TYPE "ST_CylinderHal"
VERSION : 0.1
   STRUCT
      FeedbackExtended : Bool;
      FeedbackRetracted : Bool;
      ExtendPermit : Bool;
      RetractPermit : Bool;
      PermitDiagnostic : "ST_Diagnostic";
      CoilExtend : Bool;
      CoilRetract : Bool;
   END_STRUCT;

END_TYPE

